Fanuc KAREL source: KS00026.KL

PROGRAM KS00026
%NOLOCKGROUP
TYPE
  REC_T = STRUCTURE
    VALUE: INTEGER
    FLAG: BOOLEAN
  ENDSTRUCTURE
VAR
  A: QUEUE_TYPE
  B: QUEUE_TYPE
  FLAG: BOOLEAN
  N: INTEGER
  STATUS: INTEGER
  PN: STRING[80]
  VN: STRING[80]
BEGIN
  PN = ''
  VN = 'A'
  N = ARRAY_LEN(A)
END KS00026
